(* IEC 61131-3 sources: Test-Git_ESME26/TestProgettoESME_26.fbsproj/PacDriveLib Migration/Motion/Control/Brake/FB_BrakeDisconnectionTime.fb.st^, 4 files *)

(* ---- ifBrake.prop.st ---- *)
PROPERTY ifBrake : DDI.IF_Brake
__SETTERDECLARATION__
VAR
END_VAR
__SETTERIMPLEMENTATION__
ifBrake_loc := ifBrake;

(* ---- Job.meth.st ---- *)
{attribute 'conditionalshow_all_locals'}
METHOD Job : BOOL

IF ifBrake_loc.BrakeDisconnectionTime > 0 THEN
	tBrakeDisconnectTemp := DINT_TO_TIME(ifBrake_loc.BrakeDisconnectionTime);
ELSE
	tBrakeDisconnectTemp := T#500MS;
END_IF

(* ---- timTime.prop.st ---- *)
PROPERTY INTERNAL timTime : Time
__GETTERDECLARATION__
VAR
END_VAR
__GETTERIMPLEMENTATION__
timTime:= tBrakeDisconnectTemp;

(* ---- xDone.prop.st ---- *)
PROPERTY xDone : BOOL
__GETTERDECLARATION__
VAR
END_VAR
__GETTERIMPLEMENTATION__
xDone := xDone_loc;
__SETTERDECLARATION__
VAR
END_VAR
__SETTERIMPLEMENTATION__
xDone_loc := xDone;
